(* PLC project Vn_ton_then_read, Beckhoff Automation GmbH TwinCAT PLC Control 3.5.13.21 *)
(* stored: creationDateTime 1970-01-01T00:00:00 *)

PROGRAM Vn_ton_then_read

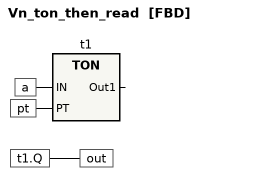
(* FBD diagram, written out as Structured Text *)
t1(IN := a, PT := pt);
out := t1.Q;
END_PROGRAM
